{attribute 'qualified_only'}
{attribute 'strict'}
TYPE E_PrLine_M_LineUsage :
(
	eNotInUse := 0,
	eMarinada_T1,
	eMarinada_T2
);
END_TYPE

(* stored: Version 1.1.0.1, ProductVersion 3.1.4024.12
   DUT E_PrLine_M_LineUsage: Id {e7844b2a-ebea-4d7e-91a5-b67c658be4f4} *)
